Staubli VAL3: insertSignal.pgx

public program insertSignal(string x_sKey, num x_nIndex, bool& x_bToSave, num x_nMoveType, num x_nActionIndex, num x_nSigValue)
  local num l_j
  local bool l_bResult
  local num l_nIndex
  local num l_i
begin
  l_nIndex=x_nIndex+1

  //insert(trajTemp:tTrajItem[x_sKey].pPointItem[l_nIndex])
  append(trajTemp:tTrajItem[x_sKey].pPointItem)

  for l_i = (size(trajTemp:tTrajItem[x_sKey].pPointItem)-1) to l_nIndex step -1
    // logMsg(toString("",l_i))
    call copyPoint3(x_sKey,l_i,l_i-1)
  endFor
  trajTemp:tTrajItem[x_sKey].pPointItem[l_nIndex].pParaItem.nMoveType=x_nMoveType

  trajTemp:tTrajItem[x_sKey].pPointItem[l_nIndex].pParaItem.nSigValue=x_nSigValue

  trajTemp:tTrajItem[x_sKey].pPointItem[l_nIndex].pParaItem.nActionIndex=x_nActionIndex



  x_bToSave=true
  //trajTemp:libSave()
end
